// TIA Portal V19 export
DATA_BLOCK "RPM"   // DB103
{ S7_Optimized_Access := 'FALSE' }
   VAR
      RAW_MIN : Array[1..20] of Int;
      RAW_MAX : Array[1..20] of Int;
      SCALE_MIN : Array[1..20] of Real;
      SCALE_MAX : Array[1..20] of Real;
      INPUT : Array[1..20] of Int;
      FAULT : Array[1..20] of Bool;
      SCALE_OUT : Array[1..20] of Real;
      STATUS : Array[1..20] of Int;
   END_VAR
BEGIN
   RAW_MAX[1..20] := 27648;
   SCALE_MAX[1..20] := 100.0;
END_DATA_BLOCK
